// TIA Portal V20 export
// export: Created 2026-11-12T08:00:00.0000000Z, ExportSetting None, DisplayName Totally Integrated Automation Portal, DisplayVersion V20, DisplayName STEP 7 Professional, DisplayVersion V20
FUNCTION_BLOCK "FB_Conveyor_BatchCounter_LAD"   // FB23, LAD
TITLE = FB_Conveyor_BatchCounter_LAD
{ S7_Optimized_Access := 'TRUE' }
// 联锁输送带与批次计数控制（严格基于 PBox + Add + Ge + Move 构建）
// stored: AutoNumber false, MemoryReserve 10, SetENOAutomatically false
   VAR_INPUT
      startCmd : Bool;
      stopCmd : Bool;
      pauseCmd : Bool;
      partSensor : Bool;
      downstreamReady : Bool;
      eStopNC : Bool;
      batchTarget : Int;
      clearCount : Bool;
   END_VAR
   VAR_OUTPUT
      conveyorRun : Bool;
      batchFull : Bool;
      partCount : Int;
   END_VAR
   VAR
      statRunning : Bool;
      statPartEdge : Bool;
      statCount : Int;
   END_VAR
   VAR_TEMP   // added for the SCL form of the ladder/FBD networks
      _w1 : Bool;
      _w2 : Bool;
   END_VAR
BEGIN

REGION Network 1: 输送带运行自锁
   // 网络1：输送带启动保持与停止/急停控制
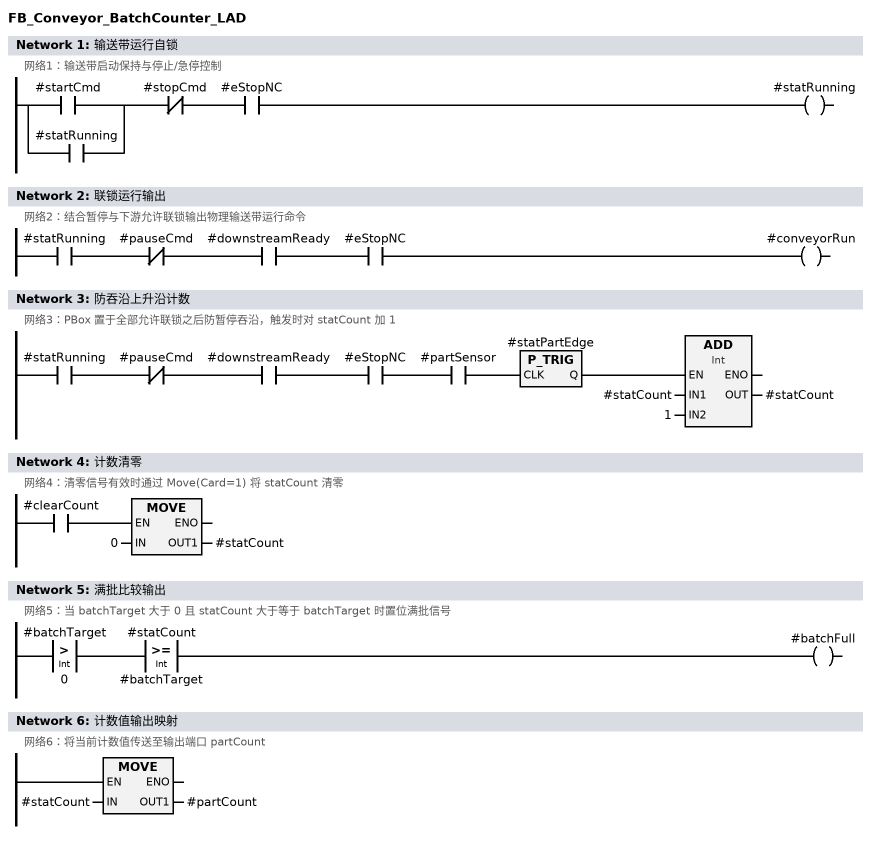
   RUNG wire#powerrail
      Contact( #startCmd )
      wire#w1
      I_Contact( #stopCmd )
      Contact( #eStopNC )
      Coil( #statRunning )
   END_RUNG
   RUNG wire#powerrail
      Contact( #statRunning )
   END_RUNG wire#w1
   // the same network as SCL:
   #statRunning := (#startCmd OR #statRunning) AND NOT #stopCmd AND #eStopNC;
END_REGION

REGION Network 2: 联锁运行输出
   // 网络2：结合暂停与下游允许联锁输出物理输送带运行命令
   RUNG wire#powerrail
      Contact( #statRunning )
      I_Contact( #pauseCmd )
      Contact( #downstreamReady )
      Contact( #eStopNC )
      Coil( #conveyorRun )
   END_RUNG
   // the same network as SCL:
   #conveyorRun := #statRunning AND NOT #pauseCmd AND #downstreamReady AND #eStopNC;
END_REGION

REGION Network 3: 防吞沿上升沿计数
   // 网络3：PBox 置于全部允许联锁之后防暂停吞沿，触发时对 statCount 加 1
   RUNG wire#powerrail
      Contact( #statRunning )
      I_Contact( #pauseCmd )
      Contact( #downstreamReady )
      Contact( #eStopNC )
      Contact( #partSensor )
      P_Trig( #statPartEdge )
      { S7_Templates := "SrcType := Int" } Add(in1 := #statCount, in2 := 1, out => #statCount)
   END_RUNG
   // the same network as SCL:
   #_w1 := #statRunning AND NOT #pauseCmd AND #downstreamReady AND #eStopNC AND #partSensor;
   #_w2 := #_w1 AND NOT #statPartEdge;   // rising edge
   #statPartEdge := #_w1;
   IF #_w2 THEN #statCount := #statCount + 1; END_IF;
END_REGION

REGION Network 4: 计数清零
   // 网络4：清零信号有效时通过 Move(Card=1) 将 statCount 清零
   RUNG wire#powerrail
      Contact( #clearCount )
      Move(in := 0, out1 => #statCount)
   END_RUNG
   // the same network as SCL:
   IF #clearCount THEN #statCount := 0; END_IF;
END_REGION

REGION Network 5: 满批比较输出
   // 网络5：当 batchTarget 大于 0 且 statCount 大于等于 batchTarget 时置位满批信号
   RUNG wire#powerrail
      { S7_Templates := "SrcType := Int" } GT_Contact(in1 := #batchTarget, in2 := 0)
      { S7_Templates := "SrcType := Int" } GE_Contact(in1 := #statCount, in2 := #batchTarget)
      Coil( #batchFull )
   END_RUNG
   // the same network as SCL:
   #batchFull := (#batchTarget > 0) AND (#statCount >= #batchTarget);
END_REGION

REGION Network 6: 计数值输出映射
   // 网络6：将当前计数值传送至输出端口 partCount
   RUNG wire#powerrail
      Move(in := #statCount, out1 => #partCount)
   END_RUNG
   // the same network as SCL:
   #partCount := #statCount;
END_REGION
END_FUNCTION_BLOCK
